RoboDK station: Car_Painting_Cell.rdk

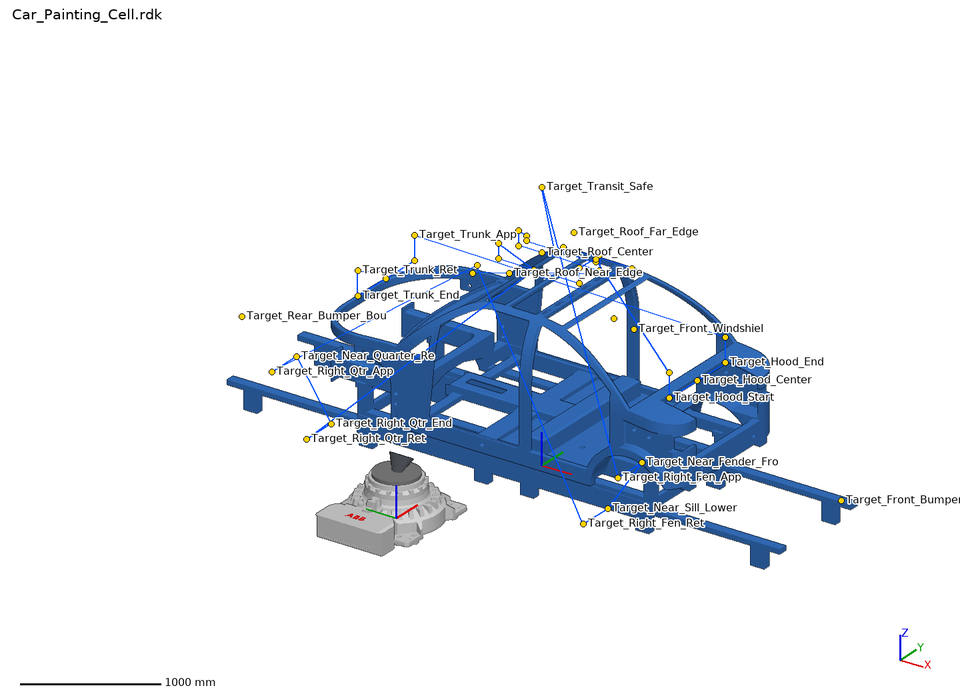
[picture v0: the station drawn from its stored meshes, robots at their saved joint values, targets as dots, program paths as lines]
Station Car_Painting_Cell (saved by RoboDK 6.0.6). Poses are relative to the parent item; angles as X-Y-Z fixed-axis rotations.
Station parameters (name, value as stored): LIN64
  - frame ABB IRB 6700-150/3.20 LeanID Base at (0, -1800, 300) mm, rotated rx 0 ry 0 rz 90 deg
    - robot ABB IRB 6700-150/3.20 LeanID: 6 axes, payload 150 kg, reach 3200 mm, repeatability 0.06 mm, weight 1280 kg
        joint limits [-170, -65, -180, -300, -130, -360] to [170, 85, 70, 300, 130, 360]; home [0, 0, 0, 0, 0, 0]; saved at [0, -10, 20, 0, 80, 180]
      - tool Paint_Gun, TCP at (0, 0, 325.06) mm, size 203.2 x 279.7 x 471.5 mm
  - frame Car_Reference_Frame at (0, 0, 0) mm
    - object Car_Body at (0, 0, 0) mm, size 4800 x 1392 x 1480 mm, geometry from Car_Body.stl
    - target Target_Roof_Center (Cartesian target) at (0, 0, 1680) mm, rotated rx 180 ry 0 rz 90 deg; joints [0, -5.605, 12.721, 0, 82.884, 180] of ABB IRB 6700-150/3.20 LeanID
    - target Target_Roof_Near_Edge (Cartesian target) at (0, -400, 1680) mm, rotated rx 180 ry 0 rz 90 deg; joints [0, -24.043, 27.41, 0, 86.633, 180] of ABB IRB 6700-150/3.20 LeanID
    - target Target_Roof_Far_Edge (Cartesian target) at (0, 400, 1680) mm, rotated rx 180 ry 0 rz 90 deg; joints [0, 12.415, -6.149, 0, 83.734, 180] of ABB IRB 6700-150/3.20 LeanID
    - target Target_Hood_Center (Cartesian target) at (1350, 0, 1050) mm, rotated rx 180 ry 0 rz 90 deg; joints [-36.87, 19.464, 8.183, 0, 62.353, 143.13] of ABB IRB 6700-150/3.20 LeanID
    - target Target_Trunk_Center (Cartesian target) at (-1350, 0, 1100) mm, rotated rx 180 ry 0 rz 90 deg; joints [36.87, 18.712, 7.248, 0, 64.04, -143.13] of ABB IRB 6700-150/3.20 LeanID
    - target Target_Front_Windshield (Cartesian target) at (800, 0, 1300) mm, rotated rx 180 ry -30 rz 180 deg; joints [-32.291, 12.078, 11.253, 25.132, 84.393, 51.256] of ABB IRB 6700-150/3.20 LeanID
    - target Target_Rear_Window (Cartesian target) at (-600, 0, 1350) mm, rotated rx 180 ry 30 rz 180 deg; joints [27.513, 7.145, 15.014, -26.507, 83.527, 124.242] of ABB IRB 6700-150/3.20 LeanID
    - target Target_Near_Fender_Front (Cartesian target) at (1500, -896, 800) mm, rotated rx 90 ry 0 rz 180 deg; joints [-81.322, 23.676, 48.283, -81.743, -87.322, 107.848] of ABB IRB 6700-150/3.20 LeanID
    - target Target_Near_Quarter_Rear (Cartesian target) at (-1500, -896, 800) mm, rotated rx 90 ry 0 rz 180 deg; joints [81.322, 23.676, 48.283, 81.743, -87.322, 72.152] of ABB IRB 6700-150/3.20 LeanID
    - target Target_Near_Sill_Lower (Cartesian target) at (1200, -896, 350) mm, rotated rx 90 ry 0 rz 180 deg; joints [-79.199, 46.895, 51.437, -79.31, -91.556, 81.813] of ABB IRB 6700-150/3.20 LeanID
    - target Target_Front_Bumper_Boundary (Cartesian target) at (2600, 0, 450) mm, rotated rx 90 ry 0 rz -90 deg; joints [-39.6, 23.445, 25.72, -39.655, -45.78, -4.095] of ABB IRB 6700-150/3.20 LeanID
    - target Target_Rear_Bumper_Boundary (Cartesian target) at (-2600, 0, 450) mm, rotated rx 90 ry 0 rz 90 deg; joints [-39.6, 23.445, 25.72, -39.655, -45.78, -4.095] of ABB IRB 6700-150/3.20 LeanID
    - target Target_Far_Side_Boundary (Cartesian target) at (0, 896, 800) mm, rotated rx 90 ry 0 rz 0 deg; joints [-39.6, 23.445, 25.72, -39.655, -45.78, -4.095] of ABB IRB 6700-150/3.20 LeanID
    - target Target_Paint_Home (joint target) at (0, -99.23, 1585.92) mm, rotated rx -180 ry 0 rz 90 deg; joints [0, -10, 20, 0, 80, 180] of ABB IRB 6700-150/3.20 LeanID
    - target Target_Roof_P1_App (Cartesian target) at (-200, -250, 1800) mm, rotated rx 180 ry 0 rz 90 deg; joints [7.352, -16.04, 17.301, 0, 88.738, 187.352] of ABB IRB 6700-150/3.20 LeanID
    - target Target_Roof_P1_Start (Cartesian target) at (-200, -250, 1680) mm, rotated rx 180 ry 0 rz 90 deg; joints [7.352, -16.403, 21.878, 0, 84.525, 187.352] of ABB IRB 6700-150/3.20 LeanID
    - target Target_Roof_P1_End (Cartesian target) at (500, -250, 1680) mm, rotated rx 180 ry 0 rz 45 deg; joints [-17.879, -13.375, 19.47, 0, 83.905, 207.121] of ABB IRB 6700-150/3.20 LeanID
    - target Target_Roof_P1_Ret (Cartesian target) at (500, -250, 1800) mm, rotated rx 180 ry 0 rz 45 deg; joints [-17.879, -13.072, 14.931, 0, 88.141, 207.121] of ABB IRB 6700-150/3.20 LeanID
    - target Target_Roof_P2_App (Cartesian target) at (500, 0, 1800) mm, rotated rx 180 ry 0 rz 45 deg; joints [-15.524, -2.357, 5.366, 0, 86.991, 209.476] of ABB IRB 6700-150/3.20 LeanID
    - target Target_Roof_P2_Start (Cartesian target) at (500, 0, 1680) mm, rotated rx 180 ry 0 rz 45 deg; joints [-15.524, -2.546, 9.835, 0, 82.711, 209.476] of ABB IRB 6700-150/3.20 LeanID
    - target Target_Roof_P2_End (Cartesian target) at (-200, 0, 1680) mm, rotated rx 180 ry 0 rz 45 deg; joints [6.34, -5.107, 12.26, 0, 82.847, 231.34] of ABB IRB 6700-150/3.20 LeanID
    - target Target_Roof_P2_Ret (Cartesian target) at (-200, 0, 1800) mm, rotated rx 180 ry 0 rz 45 deg; joints [6.34, -4.906, 7.785, 0, 87.121, 231.34] of ABB IRB 6700-150/3.20 LeanID
    - target Target_Roof_P3_App (Cartesian target) at (-200, 100, 1720) mm, rotated rx 180 ry 0 rz 45 deg; joints [6.009, -0.632, 6.536, 0, 84.096, 231.009] of ABB IRB 6700-150/3.20 LeanID
    - target Target_Roof_P3_Start (Cartesian target) at (-200, 100, 1680) mm, rotated rx 180 ry 0 rz 45 deg; joints [6.009, -0.649, 7.981, 0, 82.668, 231.009] of ABB IRB 6700-150/3.20 LeanID
    - target Target_Roof_P3_End (Cartesian target) at (400, 100, 1680) mm, rotated rx 180 ry 0 rz 45 deg; joints [-11.889, 0.745, 6.586, 0, 82.669, 213.111] of ABB IRB 6700-150/3.20 LeanID
    - target Target_Roof_P3_Ret (Cartesian target) at (400, 100, 1700) mm, rotated rx 180 ry 0 rz 45 deg; joints [-11.889, 0.748, 5.869, 0, 83.383, 213.111] of ABB IRB 6700-150/3.20 LeanID
    - target Target_Hood_App (Cartesian target) at (1350, -350, 1250) mm, rotated rx 180 ry 0 rz 0 deg; joints [-42.955, 5.144, 17.546, 0, 67.31, 227.045] of ABB IRB 6700-150/3.20 LeanID
    - target Target_Hood_Start (Cartesian target) at (1350, -350, 1050) mm, rotated rx 180 ry 0 rz 0 deg; joints [-42.955, 8.155, 21.804, 0, 60.041, 227.045] of ABB IRB 6700-150/3.20 LeanID
    - target Target_Hood_End (Cartesian target) at (1350, 350, 1050) mm, rotated rx 180 ry 0 rz 0 deg; joints [-32.125, 31.866, -8.722, 0, 66.856, 237.875] of ABB IRB 6700-150/3.20 LeanID
    - target Target_Hood_Ret (Cartesian target) at (1350, 350, 1250) mm, rotated rx 180 ry 0 rz 0 deg; joints [-32.125, 29.786, -13.094, 0, 73.308, 237.875] of ABB IRB 6700-150/3.20 LeanID
    - target Target_Trunk_App (Cartesian target) at (-1350, 350, 1300) mm, rotated rx 180 ry 0 rz 45 deg; joints [32.125, 29.424, -14.393, 0, 74.969, 257.125] of ABB IRB 6700-150/3.20 LeanID
    - target Target_Trunk_Start (Cartesian target) at (-1350, 350, 1100) mm, rotated rx 180 ry 0 rz 45 deg; joints [32.125, 31.255, -9.696, 0, 68.441, 257.125] of ABB IRB 6700-150/3.20 LeanID
    - target Target_Trunk_End (Cartesian target) at (-1350, -350, 1100) mm, rotated rx 180 ry 0 rz 45 deg; joints [42.955, 7.295, 20.84, 0, 61.865, 267.955] of ABB IRB 6700-150/3.20 LeanID
    - target Target_Trunk_Ret (Cartesian target) at (-1350, -350, 1300) mm, rotated rx 180 ry 0 rz 45 deg; joints [42.955, 4.57, 16.315, 0, 69.115, 267.955] of ABB IRB 6700-150/3.20 LeanID
    - target Target_Left_App (Cartesian target) at (400, 450, 1450) mm, rotated rx 135 ry 0 rz 0 deg; joints [-8.344, 40.786, -29.274, -7.026, 122.986, 260.24] of ABB IRB 6700-150/3.20 LeanID
    - target Target_Left_Start (Cartesian target) at (400, 550, 1450) mm, rotated rx 135 ry 0 rz 0 deg; joints [-8.053, 46.65, -38.374, -7.054, 126.232, 260.104] of ABB IRB 6700-150/3.20 LeanID
    - target Target_Left_End (Cartesian target) at (-200, 550, 1450) mm, rotated rx 135 ry 0 rz 0 deg; joints [4.046, 45.328, -36.292, 3.529, 125.842, 274.931] of ABB IRB 6700-150/3.20 LeanID
    - target Target_Left_Ret (Cartesian target) at (-200, 450, 1450) mm, rotated rx 135 ry 0 rz 0 deg; joints [4.194, 39.588, -27.458, 3.525, 122.744, 274.877] of ABB IRB 6700-150/3.20 LeanID
    - target Target_Right_Fen_App (Cartesian target) at (1500, -1200, 800) mm, rotated rx 90 ry 0 rz 180 deg; joints [-92.865, 23.284, 48.969, 87.271, 90.873, 287.726] of ABB IRB 6700-150/3.20 LeanID
    - target Target_Right_Fen_Start (Cartesian target) at (1500, -896, 800) mm, rotated rx 90 ry 0 rz 180 deg; joints [-81.322, 23.676, 48.283, 98.257, 87.322, 287.848] of ABB IRB 6700-150/3.20 LeanID
    - target Target_Right_Fen_End (Cartesian target) at (1200, -896, 350) mm, rotated rx 90 ry -45 rz 180 deg; joints [-79.199, 46.895, 51.437, 100.69, 91.556, 306.813] of ABB IRB 6700-150/3.20 LeanID
    - target Target_Right_Fen_Ret (Cartesian target) at (1200, -1200, 350) mm, rotated rx 90 ry -45 rz 180 deg; joints [-93.579, 46.927, 52.112, 86.465, 89.438, 305.978] of ABB IRB 6700-150/3.20 LeanID
    - target Target_Right_Qtr_App (Cartesian target) at (-1500, -1200, 800) mm, rotated rx 90 ry -45 rz 180 deg; joints [92.865, 23.284, 48.969, -87.271, 90.873, 297.274] of ABB IRB 6700-150/3.20 LeanID
    - target Target_Right_Qtr_Start (Cartesian target) at (-1500, -896, 800) mm, rotated rx 90 ry -45 rz 180 deg; joints [81.322, 23.676, 48.283, -98.257, 87.322, 297.152] of ABB IRB 6700-150/3.20 LeanID
    - target Target_Right_Qtr_End (Cartesian target) at (-1200, -896, 350) mm, rotated rx 90 ry 0 rz 180 deg; joints [79.199, 46.895, 51.437, -100.69, 91.556, 278.187] of ABB IRB 6700-150/3.20 LeanID
    - target Target_Right_Qtr_Ret (Cartesian target) at (-1200, -1200, 350) mm, rotated rx 90 ry 0 rz 180 deg; joints [93.579, 46.927, 52.112, -86.465, 89.438, 279.022] of ABB IRB 6700-150/3.20 LeanID
    - target Target_Transit_Safe (Cartesian target) at (0, 0, 2200) mm, rotated rx 180 ry 0 rz 0 deg; joints [0, -1.787, -9.796, 0, 101.583, 270] of ABB IRB 6700-150/3.20 LeanID
    - target Target_Transit_Right_Mid (Cartesian target) at (0, -800, 1900) mm, rotated rx 180 ry 0 rz -45 deg; joints [0, -40.798, 28.823, 0, 101.975, 315] of ABB IRB 6700-150/3.20 LeanID
  - program Car_Painting_Demo (41 instructions, listed below)
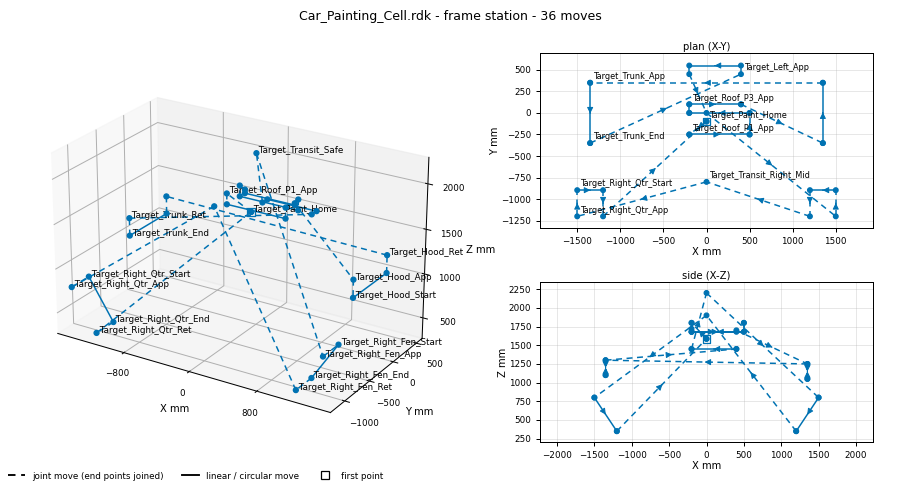
[picture p0: tool path of Car_Painting_Cell.rdk in frame station, 36 of 36 moves have a stored position in this frame; points joined in program order, loops and branches not executed]

--- program Car_Painting_Demo (robot ABB IRB 6700-150/3.20 LeanID) ---
  Set Ref.: Car_Reference_Frame
  Set Tool: Paint_Gun
  Set speed (250.0 mm/s)
  Set speed (35.0 deg/s)
  Smooth(10)
  MoveJ (Target_Paint_Home)
  MoveJ (Target_Roof_P1_App)
  MoveJ (Target_Roof_P1_Start)
  MoveL (Target_Roof_P1_End)
  MoveJ (Target_Roof_P1_Ret)
  MoveJ (Target_Roof_P2_App)
  MoveJ (Target_Roof_P2_Start)
  MoveL (Target_Roof_P2_End)
  MoveJ (Target_Roof_P2_Ret)
  MoveJ (Target_Roof_P3_App)
  MoveJ (Target_Roof_P3_Start)
  MoveL (Target_Roof_P3_End)
  MoveJ (Target_Roof_P3_Ret)
  MoveJ (Target_Hood_App)
  MoveJ (Target_Hood_Start)
  MoveL (Target_Hood_End)
  MoveJ (Target_Hood_Ret)
  MoveJ (Target_Trunk_App)
  MoveJ (Target_Trunk_Start)
  MoveL (Target_Trunk_End)
  MoveJ (Target_Trunk_Ret)
  MoveJ (Target_Left_App)
  MoveJ (Target_Left_Start)
  MoveL (Target_Left_End)
  MoveJ (Target_Left_Ret)
  MoveJ (Target_Transit_Safe)
  MoveJ (Target_Right_Fen_App)
  MoveJ (Target_Right_Fen_Start)
  MoveL (Target_Right_Fen_End)
  MoveJ (Target_Right_Fen_Ret)
  MoveJ (Target_Transit_Right_Mid)
  MoveJ (Target_Right_Qtr_App)
  MoveJ (Target_Right_Qtr_Start)
  MoveL (Target_Right_Qtr_End)
  MoveJ (Target_Right_Qtr_Ret)
  MoveJ (Target_Paint_Home)
